// TIA Portal V21 export
// export: Created 2026-11-21T13:31:41.4321747Z, ExportSetting WithDefaults, DisplayName Totally Integrated Automation Portal, DisplayVersion V21, DisplayName STEP 7 Professional, DisplayVersion V21, DisplayName STEP 7 Safety, DisplayVersion V21, DisplayName Tech WebApplication, DisplayVersion V21, DisplayName WinCC Basic/Comfort/Advanced, DisplayVersion V21, DisplayName WinCC Unified, DisplayVersion V21
VAR_GLOBAL   // PLC tag table "IO"
   Start AT %I0.0 : Bool;   // Start button
   Stop AT %I0.1 : Bool;   // Stop button
   Motor AT %Q0.0 : Bool;   // Motor contactor
   Raw AT %IW2 : Int;   // Raw level
END_VAR
